// TIA Portal V21 export
FUNCTION_BLOCK "Valve"   // FB20, LAD
TITLE = Ventil / Valve / Vanne
{ S7_Optimized_Access := 'TRUE' }
// Ein Ventil mit Rückmeldung. / A valve with feedback. / Une vanne avec retour d'information.
   VAR_INPUT
      open : Bool;   // Ventil öffnen / Open the valve / Ouvrir la vanne
      close : Bool;   // Close the valve
   END_VAR
   VAR_OUTPUT
      opened : Bool;   // Vanne ouverte
   END_VAR
   VAR
      moving : Bool;   // Ventil fährt / Valve is moving / La vanne se déplace
   END_VAR
BEGIN

REGION Network 1: Öffnen / Open / Ouvrir
   // Öffnen setzt das Fahren. / Opening starts the travel. / L'ouverture lance le déplacement.
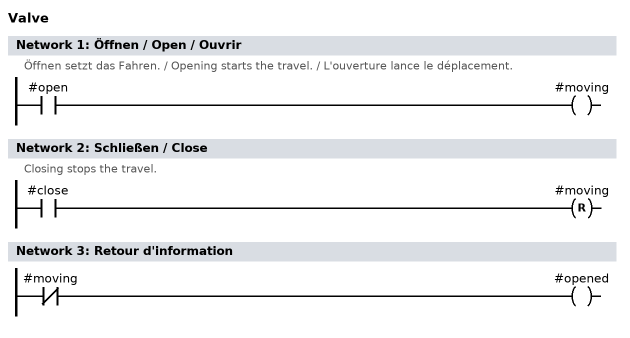
   RUNG wire#powerrail
      Contact( #open )
      Coil( #moving )
   END_RUNG
   // the same network as SCL:
   #moving := #open;
END_REGION

REGION Network 2: Schließen / Close
   // Closing stops the travel.
   RUNG wire#powerrail
      Contact( #close )
      R_Coil( #moving )
   END_RUNG
   // the same network as SCL:
   IF #close THEN #moving := FALSE; END_IF;
END_REGION

REGION Network 3: Retour d'information
   RUNG wire#powerrail
      I_Contact( #moving )
      Coil( #opened )
   END_RUNG
   // the same network as SCL:
   #opened := NOT #moving;
END_REGION
END_FUNCTION_BLOCK
